(* IEC 61131-3 sources: rusty/xtask/res (part 2) *)

(******************************************************************************
Description: Counter down
Input:
  - CD: Count down
  - LD: Load start value
  - PV: Start value
Output:
  - Q: Counter reached 0
  - CV: Current counter value
Return: Output is used as return value
***************************************************************************** *)
{external}
FUNCTION_BLOCK CTD_ULINT
VAR_INPUT
	CD : BOOL;
	LD : BOOL;
	PV : ULINT;
END_VAR
VAR_OUTPUT
	Q : BOOL;
	CV : ULINT;
END_VAR
VAR
	M : BOOL;
END_VAR
END_FUNCTION_BLOCK

(******************************************************************************
Description: Counter up and down
Input:
  - CU: Count up
  - CD: Count down
  - R: Reset counter to 0
  - LD: Load start value
  - PV: Start value / counter limit
Output:
  - QU: Counter reached limit
  - QD: Counter reached  0
  - CV: Current counter value
Return: Output is used as return value
***************************************************************************** *)
{external}
FUNCTION_BLOCK CTUD
VAR_INPUT
	CU : BOOL;
	CD : BOOL;
	R : BOOL;
	LD : BOOL;
	PV : INT;
END_VAR
VAR_OUTPUT
	QU : BOOL;
	QD : BOOL;
	CV : INT;
END_VAR
VAR
	MU : BOOL;
	MD : BOOL;
END_VAR
END_FUNCTION_BLOCK

(******************************************************************************
Description: Counter up and down
Input:
  - CU: Count up
  - CD: Count down
  - R: Reset counter to 0
  - LD: Load start value
  - PV: Start value / counter limit
Output:
  - QU: Counter reached limit
  - QD: Counter reached  0
  - CV: Current counter value
Return: Output is used as return value
***************************************************************************** *)
{external}
FUNCTION_BLOCK CTUD_INT
VAR_INPUT
	CU : BOOL;
	CD : BOOL;
	R : BOOL;
	LD : BOOL;
	PV : INT;
END_VAR
VAR_OUTPUT
	QU : BOOL;
	QD : BOOL;
	CV : INT;
END_VAR
VAR
	MU : BOOL;
	MD : BOOL;
END_VAR
END_FUNCTION_BLOCK

(******************************************************************************
Description: Counter up and down
Input:
  - CU: Count up
  - CD: Count down
  - R: Reset counter to 0
  - LD: Load start value
  - PV: Start value / counter limit
Output:
  - QU: Counter reached limit
  - QD: Counter reached  0
  - CV: Current counter value
Return: Output is used as return value
***************************************************************************** *)
{external}
FUNCTION_BLOCK CTUD_DINT
VAR_INPUT
	CU : BOOL;
	CD : BOOL;
	R : BOOL;
	LD : BOOL;
	PV : DINT;
END_VAR
VAR_OUTPUT
	QU : BOOL;
	QD : BOOL;
	CV : DINT;
END_VAR
VAR
	MU : BOOL;
	MD : BOOL;
END_VAR
END_FUNCTION_BLOCK

(******************************************************************************
Description: Counter up and down
Input:
  - CU: Count up
  - CD: Count down
  - R: Reset counter to 0
  - LD: Load start value
  - PV: Start value / counter limit
Output:
  - QU: Counter reached limit
  - QD: Counter reached  0
  - CV: Current counter value
Return: Output is used as return value
***************************************************************************** *)
{external}
FUNCTION_BLOCK CTUD_UDINT
VAR_INPUT
	CU : BOOL;
	CD : BOOL;
	R : BOOL;
	LD : BOOL;
	PV : UDINT;
END_VAR
VAR_OUTPUT
	QU : BOOL;
	QD : BOOL;
	CV : UDINT;
END_VAR
VAR
	MU : BOOL;
	MD : BOOL;
END_VAR
END_FUNCTION_BLOCK

(******************************************************************************
Description: Counter up and down
Input:
  - CU: Count up
  - CD: Count down
  - R: Reset counter to 0
  - LD: Load start value
  - PV: Start value / counter limit
Output:
  - QU: Counter reached limit
  - QD: Counter reached  0
  - CV: Current counter value
Return: Output is used as return value
***************************************************************************** *)
{external}
FUNCTION_BLOCK CTUD_LINT
VAR_INPUT
	CU : BOOL;
	CD : BOOL;
	R : BOOL;
	LD : BOOL;
	PV : LINT;
END_VAR
VAR_OUTPUT
	QU : BOOL;
	QD : BOOL;
	CV : LINT;
END_VAR
VAR
	MU : BOOL;
	MD : BOOL;
END_VAR
END_FUNCTION_BLOCK

(******************************************************************************
Description: Counter up and down
Input:
  - CU: Count up
  - CD: Count down
  - R: Reset counter to 0
  - LD: Load start value
  - PV: Start value / counter limit
Output:
  - QU: Counter reached limit
  - QD: Counter reached  0
  - CV: Current counter value
Return: Output is used as return value
***************************************************************************** *)
{external}
FUNCTION_BLOCK CTUD_ULINT
VAR_INPUT
	CU : BOOL;
	CD : BOOL;
	R : BOOL;
	LD : BOOL;
	PV : ULINT;
END_VAR
VAR_OUTPUT
	QU : BOOL;
	QD : BOOL;
	CV : ULINT;
END_VAR
VAR
	MU : BOOL;
	MD : BOOL;
END_VAR
END_FUNCTION_BLOCK (* *******************
*
* Converts little endian data format to big endian data format
*
******************** *)
{external}
FUNCTION TO_BIG_ENDIAN < T : ANY > : T
VAR_INPUT
	in : T;
END_VAR
END_FUNCTION

(********************
*
* Converts big endian data format to little endian data format
*
******************** *)
{external}
FUNCTION TO_LITTLE_ENDIAN < T : ANY > : T
VAR_INPUT
	in : T;
END_VAR
END_FUNCTION

(********************
*
* Converts to little endian data format from big endian data format
*
******************** *)
{external}
FUNCTION FROM_BIG_ENDIAN < T : ANY > : T
VAR_INPUT
	in : T;
END_VAR
END_FUNCTION

(********************
*
* Converts to big endian data format from little endian data format
*
******************** *)
{external}
FUNCTION FROM_LITTLE_ENDIAN < T : ANY > : T
VAR_INPUT
	in : T;
END_VAR
END_FUNCTION

(********************
*
* Converts LWORD to LREAL
*
******************** *)
{external}
FUNCTION LWORD_TO_LREAL : LREAL
VAR_INPUT
	in : LWORD;
END_VAR
END_FUNCTION

(********************
*
* Converts LWORD to LINT
*
******************** *)
FUNCTION LWORD_TO_LINT : LINT
VAR_INPUT
	in : LWORD;
END_VAR
	LWORD_TO_LINT := in;
END_FUNCTION

(********************
*
* Converts LWORD to DINT
*
******************** *)
FUNCTION LWORD_TO_DINT : DINT
VAR_INPUT
	in : LWORD;
END_VAR
	LWORD_TO_DINT := in;
END_FUNCTION

(********************
*
* Converts LWORD to INT
*
******************** *)
FUNCTION LWORD_TO_INT : INT
VAR_INPUT
	in : LWORD;
END_VAR
	LWORD_TO_INT := in;
END_FUNCTION

(********************
*
* Converts LWORD to SINT
*
******************** *)
FUNCTION LWORD_TO_SINT : SINT
VAR_INPUT
	in : LWORD;
END_VAR
	LWORD_TO_SINT := in;
END_FUNCTION

(********************
*
* Converts LWORD to ULINT
*
******************** *)
FUNCTION LWORD_TO_ULINT : ULINT
VAR_INPUT
	in : LWORD;
END_VAR
	LWORD_TO_ULINT := in;
END_FUNCTION

(********************
*
* Converts LWORD to UDINT
*
******************** *)
FUNCTION LWORD_TO_UDINT : UDINT
VAR_INPUT
	in : LWORD;
END_VAR
	LWORD_TO_UDINT := in;
END_FUNCTION

(********************
*
* Converts LWORD to UINT
*
******************** *)
FUNCTION LWORD_TO_UINT : UINT
VAR_INPUT
	in : LWORD;
END_VAR
	LWORD_TO_UINT := in;
END_FUNCTION

(********************
*
* Converts LWORD to USINT
*
******************** *)
FUNCTION LWORD_TO_USINT : USINT
VAR_INPUT
	in : LWORD;
END_VAR
	LWORD_TO_USINT := in;
END_FUNCTION

(********************
*
* Converts DWORD to REAL
*
******************** *)
{external}
FUNCTION DWORD_TO_REAL : REAL
VAR_INPUT
	in : DWORD;
END_VAR
END_FUNCTION

(********************
*
* Converts DWORD to LINT
*
******************** *)
FUNCTION DWORD_TO_LINT : LINT
VAR_INPUT
	in : DWORD;
END_VAR
	DWORD_TO_LINT := in;
END_FUNCTION

(********************
*
* Converts DWORD to DINT
*
******************** *)
FUNCTION DWORD_TO_DINT : DINT
VAR_INPUT
	in : DWORD;
END_VAR
	DWORD_TO_DINT := in;
END_FUNCTION

(********************
*
* Converts DWORD to INT
*
******************** *)
FUNCTION DWORD_TO_INT : INT
VAR_INPUT
	in : DWORD;
END_VAR
	DWORD_TO_INT := in;
END_FUNCTION

(********************
*
* Converts DWORD to SINT
*
******************** *)
FUNCTION DWORD_TO_SINT : SINT
VAR_INPUT
	in : DWORD;
END_VAR
	DWORD_TO_SINT := in;
END_FUNCTION

(********************
*
* Converts DWORD to ULINT
*
******************** *)
FUNCTION DWORD_TO_ULINT : ULINT
VAR_INPUT
	in : DWORD;
END_VAR
	DWORD_TO_ULINT := in;
END_FUNCTION

(********************
*
* Converts DWORD to UDINT
*
******************** *)
FUNCTION DWORD_TO_UDINT : UDINT
VAR_INPUT
	in : DWORD;
END_VAR
	DWORD_TO_UDINT := in;
END_FUNCTION

(********************
*
* Converts DWORD to UINT
*
******************** *)
FUNCTION DWORD_TO_UINT : UINT
VAR_INPUT
	in : DWORD;
END_VAR
	DWORD_TO_UINT := in;
END_FUNCTION

(********************
*
* Converts DWORD to USINT
*
******************** *)
FUNCTION DWORD_TO_USINT : USINT
VAR_INPUT
	in : DWORD;
END_VAR
	DWORD_TO_USINT := in;
END_FUNCTION

(********************
*
* Converts WORD to LINT
*
******************** *)
FUNCTION WORD_TO_LINT : LINT
VAR_INPUT
	in : WORD;
END_VAR
	WORD_TO_LINT := in;
END_FUNCTION

(********************
*
* Converts WORD to DINT
*
******************** *)
FUNCTION WORD_TO_DINT : DINT
VAR_INPUT
	in : WORD;
END_VAR
	WORD_TO_DINT := in;
END_FUNCTION

(********************
*
* Converts WORD to INT
*
******************** *)
FUNCTION WORD_TO_INT : INT
VAR_INPUT
	in : WORD;
END_VAR
	WORD_TO_INT := in;
END_FUNCTION

(********************
*
* Converts WORD to SINT
*
******************** *)
FUNCTION WORD_TO_SINT : SINT
VAR_INPUT
	in : WORD;
END_VAR
	WORD_TO_SINT := in;
END_FUNCTION

(********************
*
* Converts WORD to ULINT
*
******************** *)
FUNCTION WORD_TO_ULINT : ULINT
VAR_INPUT
	in : WORD;
END_VAR
	WORD_TO_ULINT := in;
END_FUNCTION

(********************
*
* Converts WORD to UDINT
*
******************** *)
FUNCTION WORD_TO_UDINT : UDINT
VAR_INPUT
	in : WORD;
END_VAR
	WORD_TO_UDINT := in;
END_FUNCTION

(********************
*
* Converts WORD to UINT
*
******************** *)
FUNCTION WORD_TO_UINT : UINT
VAR_INPUT
	in : WORD;
END_VAR
	WORD_TO_UINT := in;
END_FUNCTION

(********************
*
* Converts WORD to USINT
*
******************** *)
FUNCTION WORD_TO_USINT : USINT
VAR_INPUT
	in : WORD;
END_VAR
	WORD_TO_USINT := in;
END_FUNCTION

(********************
*
* Converts BYTE to LINT
*
******************** *)
FUNCTION BYTE_TO_LINT : LINT
VAR_INPUT
	in : BYTE;
END_VAR
	BYTE_TO_LINT := in;
END_FUNCTION

(********************
*
* Converts BYTE to DINT
*
******************** *)
FUNCTION BYTE_TO_DINT : DINT
VAR_INPUT
	in : BYTE;
END_VAR
	BYTE_TO_DINT := in;
END_FUNCTION

(********************
*
* Converts BYTE to INT
*
******************** *)
FUNCTION BYTE_TO_INT : INT
VAR_INPUT
	in : BYTE;
END_VAR
	BYTE_TO_INT := in;
END_FUNCTION

(********************
*
* Converts BYTE to SINT
*
******************** *)
FUNCTION BYTE_TO_SINT : SINT
VAR_INPUT
	in : BYTE;
END_VAR
	BYTE_TO_SINT := in;
END_FUNCTION

(********************
*
* Converts BYTE to ULINT
*
******************** *)
FUNCTION BYTE_TO_ULINT : ULINT
VAR_INPUT
	in : BYTE;
END_VAR
	BYTE_TO_ULINT := in;
END_FUNCTION

(********************
*
* Converts BYTE to UDINT
*
******************** *)
FUNCTION BYTE_TO_UDINT : UDINT
VAR_INPUT
	in : BYTE;
END_VAR
	BYTE_TO_UDINT := in;
END_FUNCTION

(********************
*
* Converts BYTE to UINT
*
******************** *)
FUNCTION BYTE_TO_UINT : UINT
VAR_INPUT
	in : BYTE;
END_VAR
	BYTE_TO_UINT := in;
END_FUNCTION

(********************
*
* Converts BYTE to USINT
*
******************** *)
FUNCTION BYTE_TO_USINT : USINT
VAR_INPUT
	in : BYTE;
END_VAR
	BYTE_TO_USINT := in;
END_FUNCTION

(********************
*
* Converts BOOL to LINT
*
******************** *)
FUNCTION BOOL_TO_LINT : LINT
VAR_INPUT
	in : BOOL;
END_VAR
	BOOL_TO_LINT := in;
END_FUNCTION

(********************
*
* Converts BOOL to DINT
*
******************** *)
FUNCTION BOOL_TO_DINT : DINT
VAR_INPUT
	in : BOOL;
END_VAR
	BOOL_TO_DINT := in;
END_FUNCTION

(********************
*
* Converts BOOL to INT
*
******************** *)
FUNCTION BOOL_TO_INT : INT
VAR_INPUT
	in : BOOL;
END_VAR
	BOOL_TO_INT := in;
END_FUNCTION

(********************
*
* Converts BOOL to SINT
*
******************** *)
FUNCTION BOOL_TO_SINT : SINT
VAR_INPUT
	in : BOOL;
END_VAR
	BOOL_TO_SINT := in;
END_FUNCTION

(********************
*
* Converts BOOL to ULINT
*
******************** *)
FUNCTION BOOL_TO_ULINT : ULINT
VAR_INPUT
	in : BOOL;
END_VAR
	BOOL_TO_ULINT := in;
END_FUNCTION

(********************
*
* Converts BOOL to UDINT
*
******************** *)
FUNCTION BOOL_TO_UDINT : UDINT
VAR_INPUT
	in : BOOL;
END_VAR
	BOOL_TO_UDINT := in;
END_FUNCTION

(********************
*
* Converts BOOL to UINT
*
******************** *)
FUNCTION BOOL_TO_UINT : UINT
VAR_INPUT
	in : BOOL;
END_VAR
	BOOL_TO_UINT := in;
END_FUNCTION

(********************
*
* Converts BOOL to USINT
*
******************** *)
FUNCTION BOOL_TO_USINT : USINT
VAR_INPUT
	in : BOOL;
END_VAR
	BOOL_TO_USINT := in;
END_FUNCTION

(********************
*
* Converts LREAL to LWORD
*
******************** *)
{external}
FUNCTION LREAL_TO_LWORD : LWORD
VAR_INPUT
	in : LREAL;
END_VAR
END_FUNCTION

(********************
*
* Converts REAL to DWORD
*
******************** *)
{external}
FUNCTION REAL_TO_DWORD : DWORD
VAR_INPUT
	in : REAL;
END_VAR
END_FUNCTION

(********************
*
* Converts LINT to LWORD
*
******************** *)
FUNCTION LINT_TO_LWORD : LWORD
VAR_INPUT
	in : LINT;
END_VAR
	LINT_TO_LWORD := in;
END_FUNCTION

(********************
*
* Converts LINT to DWORD
*
******************** *)
FUNCTION LINT_TO_DWORD : DWORD
VAR_INPUT
	in : LINT;
END_VAR
	LINT_TO_DWORD := in;
END_FUNCTION

(********************
*
* Converts LINT to WORD
*
******************** *)
FUNCTION LINT_TO_WORD : WORD
VAR_INPUT
	in : LINT;
END_VAR
	LINT_TO_WORD := in;
END_FUNCTION

(********************
*
* Converts LINT to BYTE
*
******************** *)
FUNCTION LINT_TO_BYTE : BYTE
VAR_INPUT
	in : LINT;
END_VAR
	LINT_TO_BYTE := in;
END_FUNCTION

(********************
*
* Converts DINT to LWORD
*
******************** *)
FUNCTION DINT_TO_LWORD : LWORD
VAR_INPUT
	in : DINT;
END_VAR
	DINT_TO_LWORD := in;
END_FUNCTION

(********************
*
* Converts DINT to DWORD
*
******************** *)
FUNCTION DINT_TO_DWORD : DWORD
VAR_INPUT
	in : DINT;
END_VAR
	DINT_TO_DWORD := in;
END_FUNCTION

(********************
*
* Converts DINT to WORD
*
******************** *)
FUNCTION DINT_TO_WORD : WORD
VAR_INPUT
	in : DINT;
END_VAR
	DINT_TO_WORD := in;
END_FUNCTION

(********************
*
* Converts DINT to BYTE
*
******************** *)
FUNCTION DINT_TO_BYTE : BYTE
VAR_INPUT
	in : DINT;
END_VAR
	DINT_TO_BYTE := in;
END_FUNCTION

(********************
*
* Converts INT to LWORD
*
******************** *)
FUNCTION INT_TO_LWORD : LWORD
VAR_INPUT
	in : INT;
END_VAR
	INT_TO_LWORD := in;
END_FUNCTION

(********************
*
* Converts INT to DWORD
*
******************** *)
FUNCTION INT_TO_DWORD : DWORD
VAR_INPUT
	in : INT;
END_VAR
	INT_TO_DWORD := in;
END_FUNCTION

(********************
*
* Converts INT to WORD
*
******************** *)
FUNCTION INT_TO_WORD : WORD
VAR_INPUT
	in : INT;
END_VAR
	INT_TO_WORD := in;
END_FUNCTION

(********************
*
* Converts INT to BYTE
*
******************** *)
FUNCTION INT_TO_BYTE : BYTE
VAR_INPUT
	in : INT;
END_VAR
	INT_TO_BYTE := in;
END_FUNCTION

(********************
*
* Converts SINT to LWORD
*
******************** *)
FUNCTION SINT_TO_LWORD : LWORD
VAR_INPUT
	in : SINT;
END_VAR
	SINT_TO_LWORD := in;
END_FUNCTION

(********************
*
* Converts SINT to DWORD
*
******************** *)
FUNCTION SINT_TO_DWORD : DWORD
VAR_INPUT
	in : SINT;
END_VAR
	SINT_TO_DWORD := in;
END_FUNCTION

(********************
*
* Converts SINT to WORD
*
******************** *)
FUNCTION SINT_TO_WORD : WORD
VAR_INPUT
	in : SINT;
END_VAR
	SINT_TO_WORD := in;
END_FUNCTION

(********************
*
* Converts SINT to BYTE
*
******************** *)
FUNCTION SINT_TO_BYTE : BYTE
VAR_INPUT
	in : SINT;
END_VAR
	SINT_TO_BYTE := in;
END_FUNCTION

(********************
*
* Converts ULINT to LWORD
*
******************** *)
FUNCTION ULINT_TO_LWORD : LWORD
VAR_INPUT
	in : ULINT;
END_VAR
	ULINT_TO_LWORD := in;
END_FUNCTION

(********************
*
* Converts ULINT to DWORD
*
******************** *)
FUNCTION ULINT_TO_DWORD : DWORD
VAR_INPUT
	in : ULINT;
END_VAR
	ULINT_TO_DWORD := in;
END_FUNCTION

(********************
*
* Converts ULINT to WORD
*
******************** *)
FUNCTION ULINT_TO_WORD : WORD
VAR_INPUT
	in : ULINT;
END_VAR
	ULINT_TO_WORD := in;
END_FUNCTION

(********************
*
* Converts ULINT to BYTE
*
******************** *)
FUNCTION ULINT_TO_BYTE : BYTE
VAR_INPUT
	in : ULINT;
END_VAR
	ULINT_TO_BYTE := in;
END_FUNCTION

(********************
*
* Converts UDINT to LWORD
*
******************** *)
FUNCTION UDINT_TO_LWORD : LWORD
VAR_INPUT
	in : UDINT;
END_VAR
	UDINT_TO_LWORD := in;
END_FUNCTION

(********************
*
* Converts UDINT to DWORD
*
******************** *)
FUNCTION UDINT_TO_DWORD : DWORD
VAR_INPUT
	in : UDINT;
END_VAR
	UDINT_TO_DWORD := in;
END_FUNCTION

(********************
*
* Converts UDINT to WORD
*
******************** *)
FUNCTION UDINT_TO_WORD : WORD
VAR_INPUT
	in : UDINT;
END_VAR
	UDINT_TO_WORD := in;
END_FUNCTION

(********************
*
* Converts UDINT to BYTE
*
******************** *)
FUNCTION UDINT_TO_BYTE : BYTE
VAR_INPUT
	in : UDINT;
END_VAR
	UDINT_TO_BYTE := in;
END_FUNCTION

(********************
*
* Converts UINT to LWORD
*
******************** *)
FUNCTION UINT_TO_LWORD : LWORD
VAR_INPUT
	in : UINT;
END_VAR
	UINT_TO_LWORD := in;
END_FUNCTION

(********************
*
* Converts UINT to DWORD
*
******************** *)
FUNCTION UINT_TO_DWORD : DWORD
VAR_INPUT
	in : UINT;
END_VAR
	UINT_TO_DWORD := in;
END_FUNCTION

(********************
*
* Converts UINT to WORD
*
******************** *)
FUNCTION UINT_TO_WORD : WORD
VAR_INPUT
	in : UINT;
END_VAR
	UINT_TO_WORD := in;
END_FUNCTION

(********************
*
* Converts UINT to BYTE
*
******************** *)
FUNCTION UINT_TO_BYTE : BYTE
VAR_INPUT
	in : UINT;
END_VAR
	UINT_TO_BYTE := in;
END_FUNCTION

(********************
*
* Converts USINT to LWORD
*
******************** *)
FUNCTION USINT_TO_LWORD : LWORD
VAR_INPUT
	in : USINT;
END_VAR
	USINT_TO_LWORD := in;
END_FUNCTION

(********************
*
* Converts USINT to DWORD
*
******************** *)
FUNCTION USINT_TO_DWORD : DWORD
VAR_INPUT
	in : USINT;
END_VAR
	USINT_TO_DWORD := in;
END_FUNCTION

(********************
*
* Converts USINT to WORD
*
******************** *)
FUNCTION USINT_TO_WORD : WORD
VAR_INPUT
	in : USINT;
END_VAR
	USINT_TO_WORD := in;
END_FUNCTION

(********************
*
* Converts USINT to BYTE
*
******************** *)
FUNCTION USINT_TO_BYTE : BYTE
VAR_INPUT
	in : USINT;
END_VAR
	USINT_TO_BYTE := in;
END_FUNCTIONVAR_GLOBAL CONSTANT
    __STRING_LENGTH : DINT := 2048;
END_VAR

(******************************************************************************
Description: String character length
Input:
    - IN:   A character string
Return: String length
***************************************************************************** *)
{external}
FUNCTION LEN < T : ANY_STRING > : DINT
VAR_INPUT {ref}
	IN : T;
END_VAR
END_FUNCTION

(******************************************************************************
Description: Left
Input:
    - IN:   A character string
    - L:    The length of the substring
Return: A substring consisting of the leftmost L characters of IN
***************************************************************************** *)
FUNCTION LEFT < T : ANY_STRING > : T
VAR_INPUT {ref}
	IN : T;
END_VAR
VAR_INPUT
    L  : DINT;
END_VAR
END_FUNCTION

{external}
FUNCTION LEFT_EXT < T : ANY_STRING > : DINT
VAR_INPUT {ref}
	IN : T;
END_VAR
VAR_INPUT
    L  : DINT;
END_VAR
VAR_IN_OUT
    OUT : T;
END_VAR
END_FUNCTION

FUNCTION LEFT__STRING : STRING[__STRING_LENGTH]
VAR_INPUT {ref}
	IN : STRING[__STRING_LENGTH];
END_VAR
VAR_INPUT
    L  : DINT;
END_VAR
    LEFT_EXT(IN, L, LEFT__STRING);
END_FUNCTION

FUNCTION LEFT__WSTRING : WSTRING[__STRING_LENGTH]
VAR_INPUT {ref}
	IN : WSTRING[__STRING_LENGTH];
END_VAR
VAR_INPUT
    L  : DINT;
END_VAR
    LEFT_EXT(IN, L, LEFT__WSTRING);
END_FUNCTION

{external}
FUNCTION LEFT_EXT__STRING : DINT
VAR_INPUT {ref}
	IN : STRING[__STRING_LENGTH];
END_VAR
VAR_INPUT
    L  : DINT;
END_VAR
VAR_IN_OUT
    OUT : STRING[__STRING_LENGTH];
END_VAR
END_FUNCTION

{external}
FUNCTION LEFT_EXT__WSTRING : DINT
VAR_INPUT {ref}
	IN : WSTRING[__STRING_LENGTH];
END_VAR
VAR_INPUT
    L  : DINT;
END_VAR
VAR_IN_OUT
    OUT : WSTRING[__STRING_LENGTH];
END_VAR
END_FUNCTION

(******************************************************************************
Description: Right
Input:
    - IN:   A character string
    - L:    The length of the substring
Return: A substring consisting of the rightmost L characters of IN
***************************************************************************** *)
FUNCTION RIGHT < T : ANY_STRING > : T
VAR_INPUT {ref}
	IN : T;
END_VAR
VAR_INPUT
    L  : DINT;
END_VAR
END_FUNCTION

{external}
FUNCTION RIGHT_EXT < T : ANY_STRING > : DINT
VAR_INPUT {ref}
	IN : T;
END_VAR
VAR_INPUT
    L  : DINT;
END_VAR
VAR_IN_OUT
    OUT : T;
END_VAR
END_FUNCTION

FUNCTION RIGHT__STRING : STRING[__STRING_LENGTH]
VAR_INPUT {ref}
	IN : STRING[__STRING_LENGTH];
END_VAR
VAR_INPUT
    L  : DINT;
END_VAR
    RIGHT_EXT(IN, L, RIGHT__STRING);
END_FUNCTION

FUNCTION RIGHT__WSTRING : WSTRING[__STRING_LENGTH]
VAR_INPUT {ref}
	IN : WSTRING[__STRING_LENGTH];
END_VAR
VAR_INPUT
    L  : DINT;
END_VAR
    RIGHT_EXT(IN, L, RIGHT__WSTRING);
END_FUNCTION

{external}
FUNCTION RIGHT_EXT__STRING : DINT
VAR_INPUT {ref}
	IN : STRING[__STRING_LENGTH];
END_VAR
VAR_INPUT
    L  : DINT;
END_VAR
VAR_IN_OUT
    OUT : STRING[__STRING_LENGTH];
END_VAR
END_FUNCTION

{external}
FUNCTION RIGHT_EXT__WSTRING : DINT
VAR_INPUT {ref}
	IN : WSTRING[__STRING_LENGTH];
END_VAR
VAR_INPUT
    L  : DINT;
END_VAR
VAR_IN_OUT
    OUT : WSTRING[__STRING_LENGTH];
END_VAR
END_FUNCTION

(******************************************************************************
Description: Middle
Input:
    - IN:   A character string
    - L:    The length of the substring
    - P:    The starting index position
Return:
    A substring that contains L characters starting
    from position P in a string.
***************************************************************************** *)
FUNCTION MID < T : ANY_STRING > : T
VAR_INPUT {ref}
	IN : T;
END_VAR
VAR_INPUT
    L  : DINT;
    P  : DINT;
END_VAR
END_FUNCTION

{external}
FUNCTION MID_EXT < T : ANY_STRING > : DINT
VAR_INPUT {ref}
	IN : T;
END_VAR
VAR_INPUT
    L  : DINT;
    P  : DINT;
END_VAR
VAR_IN_OUT
    OUT : T;
END_VAR
END_FUNCTION

FUNCTION MID__STRING : STRING[__STRING_LENGTH]
VAR_INPUT {ref}
	IN : STRING[__STRING_LENGTH];
END_VAR
VAR_INPUT
    L  : DINT;
    P  : DINT;
END_VAR
    MID_EXT(IN, L, P, MID__STRING);
END_FUNCTION

FUNCTION MID__WSTRING : WSTRING[__STRING_LENGTH]
VAR_INPUT {ref}
	IN : WSTRING[__STRING_LENGTH];
END_VAR
VAR_INPUT
    L  : DINT;
    P  : DINT;
END_VAR
    MID_EXT(IN, L, P, MID__WSTRING);
END_FUNCTION

{external}
FUNCTION MID_EXT__STRING : DINT
VAR_INPUT {ref}
	IN : STRING[__STRING_LENGTH];
END_VAR
VAR_INPUT
    L  : DINT;
    P  : DINT;
END_VAR
VAR_IN_OUT
    OUT : STRING[__STRING_LENGTH];
END_VAR
END_FUNCTION

{external}
FUNCTION MID_EXT__WSTRING : DINT
VAR_INPUT {ref}
	IN : WSTRING[__STRING_LENGTH];
END_VAR
VAR_INPUT
    L  : DINT;
    P  : DINT;
END_VAR
VAR_IN_OUT
    OUT : WSTRING[__STRING_LENGTH];
END_VAR
END_FUNCTION

(******************************************************************************
Description: Extensible concatenation
Input:
    - IN:   Two or more comma-separated strings
Return:
    A string combining all given input strings in the same order
    as the given string parameters.
***************************************************************************** *)
{external}
FUNCTION CONCAT__STRING : STRING[2048]
VAR_INPUT {ref}
	args : {sized} STRING...;
END_VAR
END_FUNCTION

{external}
FUNCTION CONCAT__WSTRING : WSTRING[2048]
VAR_INPUT {ref}
	args : {sized} WSTRING...;
END_VAR
END_FUNCTION

FUNCTION CONCAT < T : ANY_STRING > : T
VAR_INPUT {ref}
	args : {sized} T...;
END_VAR
END_FUNCTION

{external}
FUNCTION CONCAT_EXT < T : ANY_STRING > : DINT
VAR_IN_OUT
    OUT : T;
END_VAR
VAR_INPUT {ref}
    args : {sized} T...;
END_VAR
END_FUNCTION

(******************************************************************************
Description: Insert
Input:
    IN1:    The string to insert into
    IN2:    The string to insert
    P:      The position at which to insert
Return:
    A string consisting of IN2 inserted at position P into string IN1
***************************************************************************** *)
FUNCTION INSERT < T : ANY_STRING > : T
VAR_INPUT {ref}
	IN1 : T;
    IN2 : T;
END_VAR
VAR_INPUT
    P   : DINT;
END_VAR
END_FUNCTION

{external}
FUNCTION INSERT_EXT < T : ANY_STRING > : DINT
VAR_INPUT {ref}
	IN1 : T;
    IN2 : T;
END_VAR
VAR_INPUT
    P   : DINT;
END_VAR
VAR_IN_OUT
    OUT : T;
END_VAR
END_FUNCTION

FUNCTION INSERT__STRING : STRING[__STRING_LENGTH]
VAR_INPUT {ref}
	IN1 : STRING[__STRING_LENGTH];
    IN2 : STRING[__STRING_LENGTH];
END_VAR
VAR_INPUT
    P   : DINT;
END_VAR
    INSERT_EXT(IN1, IN2, P, INSERT__STRING);
END_FUNCTION

FUNCTION INSERT__WSTRING : WSTRING[__STRING_LENGTH]
VAR_INPUT {ref}
	IN1 : WSTRING[__STRING_LENGTH];
    IN2 : WSTRING[__STRING_LENGTH];
END_VAR
VAR_INPUT
    P   : DINT;
END_VAR
    INSERT_EXT(IN1, IN2, P, INSERT__WSTRING);
END_FUNCTION

{external}
FUNCTION INSERT_EXT__STRING : DINT
VAR_INPUT {ref}
	IN1 : STRING[__STRING_LENGTH];
    IN2 : STRING[__STRING_LENGTH];
END_VAR
VAR_INPUT
    P   : DINT;
END_VAR
VAR_IN_OUT
    OUT : STRING[__STRING_LENGTH];
END_VAR
END_FUNCTION

{external}
FUNCTION INSERT_EXT__WSTRING : DINT
VAR_INPUT {ref}
	IN1 : WSTRING[__STRING_LENGTH];
    IN2 : WSTRING[__STRING_LENGTH];
END_VAR
VAR_INPUT
    P   : DINT;
END_VAR
VAR_IN_OUT
    OUT : WSTRING[__STRING_LENGTH];
END_VAR
END_FUNCTION

(******************************************************************************
Description: Delete
Input:
    IN: The string to delete characters from
    L:  The amount of characters to delete
    P:  The position at which to start deleting
Return: A new string with L characters deleted from P onwards
***************************************************************************** *)
FUNCTION DELETE < T : ANY_STRING > : T
VAR_INPUT {ref}
	IN : T;
END_VAR
VAR_INPUT
    L  : DINT;
    P  : DINT;
END_VAR
END_FUNCTION

{external}
FUNCTION DELETE_EXT < T : ANY_STRING > : DINT
VAR_INPUT {ref}
	IN : T;
END_VAR
VAR_INPUT
    L  : DINT;
    P  : DINT;
END_VAR
VAR_IN_OUT
    OUT : T;
END_VAR
END_FUNCTION

FUNCTION DELETE__STRING : STRING[__STRING_LENGTH]
VAR_INPUT {ref}
	IN : STRING[__STRING_LENGTH];
END_VAR
VAR_INPUT
    L  : DINT;
    P  : DINT;
END_VAR
    DELETE_EXT(IN, L, P, DELETE__STRING);
END_FUNCTION

FUNCTION DELETE__WSTRING : WSTRING[__STRING_LENGTH]
VAR_INPUT {ref}
	IN : WSTRING[__STRING_LENGTH];
END_VAR
VAR_INPUT
    L  : DINT;
    P  : DINT;
END_VAR
    DELETE_EXT(IN, L, P, DELETE__WSTRING);
END_FUNCTION

{external}
FUNCTION DELETE_EXT__STRING : DINT
VAR_INPUT {ref}
	IN : STRING[__STRING_LENGTH];
END_VAR
VAR_INPUT
    L  : DINT;
    P  : DINT;
END_VAR
VAR_IN_OUT
    OUT : STRING[__STRING_LENGTH];
END_VAR
END_FUNCTION

{external}
FUNCTION DELETE_EXT__WSTRING : DINT
VAR_INPUT {ref}
	IN : WSTRING[__STRING_LENGTH];
END_VAR
VAR_INPUT
    L  : DINT;
    P  : DINT;
END_VAR
VAR_IN_OUT
    OUT : WSTRING[__STRING_LENGTH];
END_VAR
END_FUNCTION
(******************************************************************************
Description: Replace
Input:
    IN1:    The string to replace characters from
    IN2:    The replacement string to be inserted
    L:      The amount of characters to delete
    P:      The position at which to start deleting
Return: A new string which has L characters replaced by IN2 from position P onwards
***************************************************************************** *)
FUNCTION REPLACE < T : ANY_STRING > : T
VAR_INPUT {ref}
	IN1 : T;
    IN2 : T;
END_VAR
VAR_INPUT
    L  : DINT;
    P  : DINT;
END_VAR
END_FUNCTION

{external}
FUNCTION REPLACE_EXT < T : ANY_STRING > : DINT
VAR_INPUT {ref}
    IN1 : T;
    IN2 : T;
END_VAR
VAR_INPUT
    L   : DINT;
    P   : DINT;
END_VAR
VAR_IN_OUT
    OUT : T;
END_VAR
END_FUNCTION

FUNCTION REPLACE__STRING : STRING[__STRING_LENGTH]
VAR_INPUT {ref}
	IN1 : STRING[__STRING_LENGTH];
    IN2 : STRING[__STRING_LENGTH];
END_VAR
VAR_INPUT
    L  : DINT;
    P  : DINT;
END_VAR
    REPLACE_EXT(IN1, IN2, L, P, REPLACE__STRING);
END_FUNCTION

FUNCTION REPLACE__WSTRING : WSTRING[__STRING_LENGTH]
VAR_INPUT {ref}
    IN1 : WSTRING[__STRING_LENGTH];
    IN2 : WSTRING[__STRING_LENGTH];
END_VAR
VAR_INPUT
    L   : DINT;
    P   : DINT;
END_VAR
    REPLACE_EXT(IN1, IN2, L, P, REPLACE__WSTRING);
END_FUNCTION

{external}
FUNCTION REPLACE_EXT__STRING : DINT
VAR_INPUT {ref}
    IN1 : STRING[__STRING_LENGTH];
    IN2 : STRING[__STRING_LENGTH];
END_VAR
VAR_INPUT
    L   : DINT;
    P   : DINT;
END_VAR
VAR_IN_OUT
    OUT : STRING[__STRING_LENGTH];
END_VAR
END_FUNCTION

{external}
FUNCTION REPLACE_EXT__WSTRING : DINT
VAR_INPUT {ref}
    IN1 : WSTRING[__STRING_LENGTH];
    IN2 : WSTRING[__STRING_LENGTH];
END_VAR
VAR_INPUT
    L   : DINT;
    P   : DINT;
END_VAR
VAR_IN_OUT
    OUT : WSTRING[__STRING_LENGTH];
END_VAR
END_FUNCTION

(******************************************************************************
Description: Find
Input:
    IN1:    The string in which to search in
    IN2:    The substring to search for
Return: The character index of the first match. 0 if there are no matches.
***************************************************************************** *)
{external}
FUNCTION FIND < T : ANY_STRING > : DINT
VAR_INPUT {ref}
	IN1 : T;
    IN2 : T;
END_VAR
END_FUNCTION

(******************************************************************************
Description: Decreasing sequence
Input:  The strings to compare, in order. ((IN1>IN2) & (IN2>IN3) & .. & (INn-1>INn))
Return:
    TRUE if codepoints are in decreasing order (alphabetical order: ZYX > YXW > XWV ..)
    FALSE otherwise
***************************************************************************** *)
{external}
FUNCTION GT < T : ANY_STRING > : BOOL
VAR_INPUT {ref}
	IN1 : {sized} T...;
END_VAR
END_FUNCTION

// passing strings by ref causes an error/warning. code still compiles and works correctly
FUNCTION STRING_GREATER : BOOL
VAR_INPUT
    a, b : STRING;
END_VAR
    STRING_GREATER := GT(a, b);
END_FUNCTION

FUNCTION WSTRING_GREATER : BOOL
VAR_INPUT
    a, b : WSTRING;
END_VAR
    WSTRING_GREATER := GT(a, b);
END_FUNCTION
(******************************************************************************
Description: Monotonic sequence
Input:  The strings to compare, in order. ((IN1>=IN2) & (IN2>=IN3) & .. & (INn-1>=INn))
Return:
    TRUE if codepoints are in decreasing order or are equal to adjacent codepoints (alphabetical order: ZYX >= ZYX >= YXW ..)
    FALSE otherwise
***************************************************************************** *)
{external}
FUNCTION GE < T : ANY_STRING > : BOOL
VAR_INPUT {ref}
	IN1 : {sized} T...;
END_VAR
END_FUNCTION

(******************************************************************************
Description: Equality
Input: The strings to compare, in order. ((IN1=IN2) & (IN2=IN3) & .. & (INn-1=INn))
Return:
    TRUE if codepoints are equal to each other
    FALSE otherwise.
***************************************************************************** *)
{external}
FUNCTION EQ < T : ANY_STRING > : BOOL
VAR_INPUT {ref}
	IN1 : {sized} T...;
END_VAR
END_FUNCTION

FUNCTION STRING_EQUAL : BOOL
VAR_INPUT
    a, b : STRING;
END_VAR
    STRING_EQUAL := EQ(a, b);
END_FUNCTION

FUNCTION WSTRING_EQUAL : BOOL
VAR_INPUT
    a, b : WSTRING;
END_VAR
    WSTRING_EQUAL := EQ(a, b);
END_FUNCTION

(******************************************************************************
Description: Monotonic sequence
Input:  The strings to compare, in order. ((IN1<=IN2) & (IN2<=IN3) & .. & (INn-1<=INn))
Return:
    TRUE if codepoints are in increasing order or are equal to adjacent codepoints (alphabetical order: ABC <= ABC <= BCD ..)
    FALSE otherwise
***************************************************************************** *)
{external}
FUNCTION LE < T : ANY_STRING > : BOOL
VAR_INPUT {ref}
	IN1 : {sized} T...;
END_VAR
END_FUNCTION

(******************************************************************************
Description: Increasing sequence
Input:  The strings to compare, in order. ((IN1<IN2) & (IN2<IN3) & .. & (INn-1<INn))
Return:
    TRUE if codepoints are in increasing order (alphabetical order: ABC < BCD < CDE ..)
    FALSE otherwise
***************************************************************************** *)
{external}
FUNCTION LT < T : ANY_STRING > : BOOL
VAR_INPUT {ref}
	IN1 : {sized} T...;
END_VAR
END_FUNCTION

FUNCTION STRING_LESS : BOOL
VAR_INPUT
    a, b : STRING;
END_VAR
    STRING_LESS := LT(a, b);
END_FUNCTION

FUNCTION WSTRING_LESS : BOOL
VAR_INPUT
    a, b : WSTRING;
END_VAR
    WSTRING_LESS := LT(a, b);
END_FUNCTION

(******************************************************************************
Description: Inequality
Input: The strings to compare. (IN1<>IN2)
Return:
    TRUE if strings do not match
    FALSE otherwise
***************************************************************************** *)
{external}
FUNCTION NE < T : ANY_STRING > : BOOL
VAR_INPUT {ref}
	IN1 : T;
    IN2 : T;
END_VAR
END_FUNCTION (* Definitions of arithmetic functions defined by the IEC61131-3 standard *)

{external}
VAR_GLOBAL
	PI_REAL : REAL;
	PI_LREAL : LREAL;
	FRAC_PI_2_REAL : REAL;
	FRAC_PI_2_LREAL : LREAL;
	FRAC_PI_4_REAL : REAL;
	FRAC_PI_4_LREAL : LREAL;
	E_REAL : REAL;
	E_LREAL : LREAL;
END_VAR

(* Calculates the square root of a given value *)
{external}
FUNCTION SQRT < T : ANY_REAL > : T
VAR_INPUT
	in : T;
END_VAR
END_FUNCTION

(** Logarithmic functions * *)

(* Calculates the natural logarithm of the given value *)
{external}
FUNCTION LN < T : ANY_REAL > : T
VAR_INPUT
	in : T;
END_VAR
END_FUNCTION

(* Calculates the base 10 logarithm of the given value *)
{external}
FUNCTION LOG < T : ANY_REAL > : T
VAR_INPUT
	in : T;
END_VAR
END_FUNCTION

(* Calculates the natural exporenent of the given value *)
{external}
FUNCTION EXP < T : ANY_REAL > : T
VAR_INPUT
	in : T;
END_VAR
END_FUNCTION

(** Trigonometric functions * *)

(* Calculates the sine of the given value in radiants *)
{external}
FUNCTION SIN < T : ANY_REAL > : T
VAR_INPUT
	rad : T;
END_VAR
END_FUNCTION

(* Calculates the cosine of the given value in radiants *)
{external}
FUNCTION COS < T : ANY_REAL > : T
VAR_INPUT
	rad : T;
END_VAR
END_FUNCTION

(* Calculates the tangent of the given value in radiants *)
{external}
FUNCTION TAN < T : ANY_REAL > : T
VAR_INPUT
	rad : T;
END_VAR
END_FUNCTION

(* Calculates the arc sine of the given value *)
{external}
FUNCTION ASIN < T : ANY_REAL > : T
VAR_INPUT
	in : T;
END_VAR
END_FUNCTION

(* Calculates the arc cosine of the given value *)
{external}
FUNCTION ACOS < T : ANY_REAL > : T
VAR_INPUT
	in : T;
END_VAR
END_FUNCTION

(* Calculates the arc tangent of the given value *)
{external}
FUNCTION ATAN < T : ANY_REAL > : T
VAR_INPUT
	in : T;
END_VAR
END_FUNCTION

(* Calculate the four quadrant arc tangent of the given values *)
{external}
FUNCTION ATAN2 < T : ANY_REAL > : T
VAR_INPUT
	y : T;
	x : T;
END_VAR
END_FUNCTION

{external}
FUNCTION EXPT < T : ANY_REAL, U : ANY_NUM > : T
VAR_INPUT
	in1 : T;
	in2 : U;
END_VAR
END_FUNCTION

{external}
FUNCTION EXPT__REAL__DINT : REAL
VAR_INPUT
	in1 : REAL;
	in2 : DINT;
END_VAR
END_FUNCTION

{external}
FUNCTION EXPT__REAL__REAL : REAL
VAR_INPUT
	in1 : REAL;
	in2 : REAL;
END_VAR
END_FUNCTION

(* LREAL to REAL conversion will happen for the exponent
   This will produce the closest possible REAL value
   On overflow, infinity of the same sign as the input is produced *)
{external}
FUNCTION EXPT__REAL__LREAL : REAL
VAR_INPUT
	in1 : REAL;
	in2 : LREAL;
END_VAR
END_FUNCTION

{external}
FUNCTION EXPT__LREAL__DINT : LREAL
VAR_INPUT
	in1 : LREAL;
	in2 : DINT;
END_VAR
END_FUNCTION

{external}
FUNCTION EXPT__LREAL__REAL : LREAL
VAR_INPUT
	in1 : LREAL;
	in2 : REAL;
END_VAR
END_FUNCTION

{external}
FUNCTION EXPT__LREAL__LREAL : LREAL
VAR_INPUT
	in1 : LREAL;
	in2 : LREAL;
END_VAR
END_FUNCTION

FUNCTION EXPT__REAL__USINT : REAL
VAR_INPUT
	in1 : REAL;
	in2 : USINT;
END_VAR
    EXPT__REAL__USINT := EXPT__REAL__DINT(in1, in2);
END_FUNCTION

FUNCTION EXPT__REAL__UINT : REAL
VAR_INPUT
	in1 : REAL;
	in2 : UINT;
END_VAR
    EXPT__REAL__UINT := EXPT__REAL__DINT(in1, in2);
END_FUNCTION

FUNCTION EXPT__REAL__UDINT : REAL
VAR_INPUT
	in1 : REAL;
	in2 : UDINT;
END_VAR
    EXPT__REAL__UDINT := EXPT__REAL__DINT(in1, in2);
END_FUNCTION

FUNCTION EXPT__REAL__ULINT : REAL
VAR_INPUT
	in1 : REAL;
	in2 : ULINT;
END_VAR
    EXPT__REAL__ULINT := EXPT__REAL__DINT(in1, in2);
END_FUNCTION

FUNCTION EXPT__REAL__SINT : REAL
VAR_INPUT
	in1 : REAL;
	in2 : SINT;
END_VAR
    EXPT__REAL__SINT := EXPT__REAL__DINT(in1, in2);
END_FUNCTION

FUNCTION EXPT__REAL__INT : REAL
VAR_INPUT
	in1 : REAL;
	in2 : INT;
END_VAR
    EXPT__REAL__INT := EXPT__REAL__DINT(in1, in2);
END_FUNCTION

FUNCTION EXPT__REAL__LINT : REAL
VAR_INPUT
	in1 : REAL;
	in2 : LINT;
END_VAR
    EXPT__REAL__LINT := EXPT__REAL__DINT(in1, in2);
END_FUNCTION

FUNCTION EXPT__LREAL__USINT : LREAL
VAR_INPUT
	in1 : LREAL;
	in2 : USINT;
END_VAR
    EXPT__LREAL__USINT := EXPT__LREAL__DINT(in1, in2);
END_FUNCTION

FUNCTION EXPT__LREAL__UINT : LREAL
VAR_INPUT
	in1 : LREAL;
	in2 : UINT;
END_VAR
    EXPT__LREAL__UINT := EXPT__LREAL__DINT(in1, in2);
END_FUNCTION

FUNCTION EXPT__LREAL__UDINT : LREAL
VAR_INPUT
	in1 : LREAL;
	in2 : UDINT;
END_VAR
    EXPT__LREAL__UDINT := EXPT__LREAL__DINT(in1, in2);
END_FUNCTION

FUNCTION EXPT__LREAL__ULINT : LREAL
VAR_INPUT
	in1 : LREAL;
	in2 : ULINT;
END_VAR
    EXPT__LREAL__ULINT := EXPT__LREAL__DINT(in1, in2);
END_FUNCTION

FUNCTION EXPT__LREAL__SINT : LREAL
VAR_INPUT
	in1 : LREAL;
	in2 : SINT;
END_VAR
    EXPT__LREAL__SINT := EXPT__LREAL__DINT(in1, in2);
END_FUNCTION

FUNCTION EXPT__LREAL__INT : LREAL
VAR_INPUT
	in1 : LREAL;
	in2 : INT;
END_VAR
    EXPT__LREAL__INT := EXPT__LREAL__DINT(in1, in2);
END_FUNCTION

FUNCTION EXPT__LREAL__LINT : LREAL
VAR_INPUT
	in1 : LREAL;
	in2 : LINT;
END_VAR
    EXPT__LREAL__LINT := EXPT__LREAL__DINT(in1, in2);
END_FUNCTION
(**************************
 *
 *This operator returns the absolute value of a number.
 *
************************ *)
FUNCTION ABS < T : ANY_NUM > : T
VAR_INPUT
	IN : T;
END_VAR

END_FUNCTION

(* Specialized implementation of ABS for DINT *)
/* FUNCTION ABS__DINT : DINT */
FUNCTION ABS__DINT : DINT
VAR_INPUT
	IN : DINT;
END_VAR
	ABS__DINT := IN;
	IF ABS__DINT < 0 THEN
		ABS__DINT := - 1 * ABS__DINT;
	END_IF
END_FUNCTION

(* Specialized implementation of ABS for SINT *)
FUNCTION ABS__SINT : SINT
VAR_INPUT
	IN : SINT;
END_VAR
	ABS__SINT := ABS__DINT(IN);
END_FUNCTION

(* Specialized implementation of ABS for INT *)
FUNCTION ABS__INT : INT
VAR_INPUT
	IN : INT;
END_VAR
	ABS__INT := ABS__DINT(IN);
END_FUNCTION

(* Specialized implementation of ABS for LINT *)
FUNCTION ABS__LINT : LINT
VAR_INPUT
	IN : LINT;
END_VAR
	ABS__LINT := IN;
	IF ABS__LINT < 0 THEN
		ABS__LINT := - 1 * ABS__LINT;
	END_IF
END_FUNCTION

(* Specialized implementation of ABS for REAL *)
FUNCTION ABS__REAL : REAL
VAR_INPUT
	IN : REAL;
END_VAR
	ABS__REAL := ABS__LREAL(IN);
END_FUNCTION

(* Specialized implementation of ABS for LREAL *)
FUNCTION ABS__LREAL : LREAL
VAR_INPUT
	IN : LREAL;
END_VAR
	ABS__LREAL := IN;
	IF ABS__LREAL < 0 THEN
		ABS__LREAL := - 1.0 * ABS__LREAL;
	END_IF
END_FUNCTION

(**************************
 *
 * Rounds a given ANY_REAL to the nearest integer
 * Rounds half values away from zero
 *
************************ *)
{external}
FUNCTION ROUND < T : ANY_REAL > : T
VAR_INPUT
	in : T;
END_VAR
END_FUNCTION
CLASS MyClass
    VAR
        x, y : INT;
    END_VAR

    METHOD testMethod
        VAR_INPUT myMethodArg : INT; END_VAR
        VAR myMethodLocalVar : INT; END_VAR

        x := myMethodArg;
    END_METHOD
END_CLASSPROGRAM name
(1 + 2) * (3 + 4);
END_PROGRAM
FUNCTION smaller_than_ten : BOOL
	VAR_INPUT
		n : INT;
	END_VAR

	IF n < 10 THEN
		smaller_than_ten := TRUE;
		RETURN;
	END_IF;
	smaller_than_ten := FALSE;
END_FUNCTION
PROGRAM hello
VAR
   x : INT
   y : BOOL;
END_VAR
   IF x = 2 THEN
      x := 3
END_PROGRAM
FUNCTION a : DINT END_FUNCTION
        PROGRAM main
        VAR
            x : ARRAY[0..1] OF INT;
            y : REF_TO INT;
            z : REF_TO ARRAY[0..1] OF INT;
        END_VAR
            x[0] := 1;
            y^ := 2;
            y^.1 := 3;
            z^[0] := 4;
            z^[1].1 := 5;
						a() := 5;
        END_PROGRAM
@EXTERNAL FUNCTION LOG : DINT
VAR_INPUT
    x : DINT;
END_VAR
END_FUNCTION

@EXTERNAL FUNCTION PRINTF : DINT
VAR_INPUT
    text : STRING;
    value : DINT;
END_VAR
END_FUNCTION

FUNCTION main : DINT
	main := LOG(100);
  PRINTF('Log value %d\n', main);
END_FUNCTION
FUNCTION main : DINT
  main := 1;
  WHILE main < 10 DO
    main := main + 1;
    CONTINUE;
    main := 200;
  END_WHILE
END_FUNCTION
TYPE MyStruct : STRUCT  x : DINT; y : DINT; END_STRUCT END_TYPE

FUNCTION main : DINT
	main := foo();
END_FUNCTION

FUNCTION foo : DINT
VAR
				x : DINT;
				s : MyStruct;
				u, y : REF_TO DINT;
				z : REF_TO REF_TO DINT;

END_VAR
u := NULL;
u := &s.x;
y := u;
z := &y;
s.x := 9;
z^^ := y^ * 2;
y^ := z^^ * 2;

foo := y^;
END_FUNCTION
{external}
FUNCTION puts : DINT
VAR_INPUT {ref}
    text : STRING;
END_VAR
END_FUNCTION

FUNCTION main : DINT
	puts('hello, world!$N');
END_FUNCTION
PROGRAM hello
VAR
   x : INT;
   y : INT;
   z : INT;
END_VAR

IF Condition THEN

ELSIF

END_IF;

1 + 2 + 3 + 4;
END_PROGRAM
PROGRAM exp a AND NOT b OR c XOR d; END_PROGRAMPROGRAM prg
    VAR
			a : INT;
			b : REAL;
    END_VAR
		b := 1.5;
		a := b;
END_PROGRAM
PROGRAM a
(* C�mment *)
END_PROGRAM
PROGRAM a
    VAR
        binvar      AT %IX7.8 : BOOL;
        sinvar      AT %IB4.8 : BYTE;
        winvar      AT %IW3.1 : WORD;
        dinvar      AT %ID1.7 : DWORD;
        boutvar     AT %QX7.7 : BOOL;
        soutvar     AT %QB1.6 : BYTE;
        woutvar     AT %QW2.4 : WORD;
        doutvar     AT %QD1.4 : DWORD;
        bmemvar     AT %MX7.8 : BOOL;
        smemvar     AT %MB5.8 : BYTE;
        wmemvar     AT %MW4.2 : WORD;
        dmemvar     AT %MD8.3 : DWORD;
        linvar      AT %IL9.0 : LWORD;
        loutvar     AT %QL4.2 : LWORD;
        lmemvar     AT %ML9.6 : LWORD;
    END_VAR
END_PROGRAM
PROGRAM a
(* Cömment *)
END_PROGRAM
FUNCTION myFunc : DINT
VAR_INPUT
	 a, b, c : DINT;
END_VAR
END_FUNCTION
FUNCTION foo2 : LINT
    foo2 := CONCAT_DATE(INT#4, SINT#5, SINT#6);
END_FUNCTION{external}
FUNCTION CONCAT_DATE < T : ANY_INT > : DATE
VAR_INPUT
	year : T;
	month : T;
	day : T;
END_VAR
END_FUNCTION

FUNCTION main : INT
VAR_INPUT

END_VAR

VAR

END_VAR
mainProg();
main := mainProg.a;

END_FUNCTION
PROGRAM mainProg
VAR
	a : DINT := 0;
END_VAR
a := 42;
END_PROGRAM
FUNCTION foo1 : LINT
    foo1 := CONCAT_DATE(INT#1, SINT#2, SINT#3);
END_FUNCTIONVAR_GLOBAL CONSTANT
	myValue : BOOL := TRUE;
END_VAR

FUNCTION_BLOCK myFb2
	VAR
		fb : myFb;
	END_VAR
END_FUNCTION_BLOCK
VAR_GLOBAL CONSTANT
	myValue2 : BOOL := TRUE;
END_VAR

VAR_GLOBAL CONSTANT
	myValue : BOOL := TRUE;
END_VAR

FUNCTION_BLOCK myFB
	VAR
		myS : myStruct := (a := 2);
	END_VAR
END_FUNCTION_BLOCK
{external}
FUNCTION func1 : DINT
END_FUNCTION

FUNCTION func2 : DINT
	func1();
END_FUNCTION

FUNCTION relative : DINT
END_FUNCTION
TYPE myStruct : STRUCT
	a : INT := 5;
	b : DINT := 6;
END_STRUCT
END_TYPE
{external}
FUNCTION func2 : DINT
END_FUNCTION

FUNCTION func1 : DINT
	func2();
END_FUNCTION

PROGRAM name
(1 + 2) * (3 + 4);
END_PROGRAM
PROGRAM hello
VAR
   x : INT;
   y : BOOL;
END_VAR
   IF x = 2 THEN
      x := 3;
   END_IF
END_PROGRAM
PROGRAM prg
    VAR
			a : INT;
			b : REAL;
    END_VAR
		b := 1.5;
		a := b;
END_PROGRAM
VAR_GLOBAL
    flags : ARRAY[1..500_000_000] OF BOOL;
    sieve_size : ULINT := 500_000_000;
END_VAR

// en.wikipedia.org/wiki/Sieve_of_Eratosthenes
FUNCTION sieve : DINT
    VAR
        i, j : ULINT;
        primes : ULINT;
    END_VAR

    FOR i := 2 TO sieve_size DO
        IF flags[i] = 0 THEN
            FOR j := i * i TO sieve_size BY i DO
                IF j < sieve_size THEN
                    flags[j] := 1;
                END_IF;
            END_FOR;
        END_IF;
    END_FOR;

    FOR i := 2 TO sieve_size DO
        IF flags[i] = 0 THEN
            primes := primes + 1;
        END_IF;
    END_FOR;

    printf('Primes found: %lld (correct: %d)$N', primes, (primes - 1) = 26_355_867);
END_FUNCTION

FUNCTION main : DINT
    sieve();
END_FUNCTION

{external}
FUNCTION printf : DINT
    VAR_INPUT {ref} format : STRING; END_VAR
    VAR_INPUT args : ...; END_VAR
END_FUNCTIONTYPE struct2 :
STRUCT
    param1 : DINT;
    param2 : DINT;
END_STRUCT
END_TYPE

PROGRAM mainProg
    VAR
        node : ARRAY[0..15] OF struc2 := ((param1 := 1, param2 := 2), (param1 := 3, param2 := 4));
        // node : ARRAY[0..15] OF struct2 := [(param1 := 1, param2 := 2), (param1 := 3, param2 := 4)];
    END_VAR
END_PROGRAM
